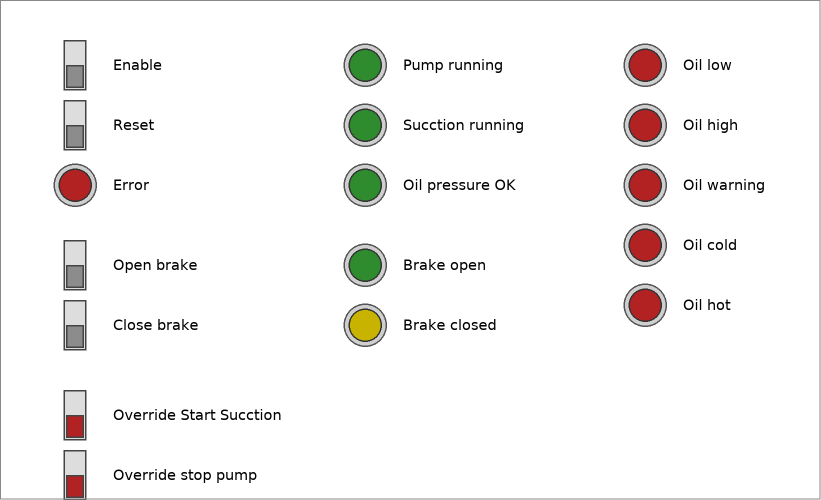
VISUALIZATION Hydraulics  // 821x500
    DipSwitch (50,40 50x50), variable: HydraulicsControl.enable, behaviour: TOGGLE, style: Switch-DipSwitch-Gray
    DipSwitch (50,100 50x50), variable: HydraulicsControl.reset, behaviour: TOGGLE, style: Switch-DipSwitch-Gray
    Label (110,50 101x30), "Enable"
    Label (110,110 101x30), "Reset"
    Lamp1 (50,160 50x50), variable: HydraulicsControl.error, style: Lamp-Lamp1-Red
    Label (110,170 101x30), "Error"
    DipSwitch (50,390 50x50), variable: HydraulicsControl.suction_manual, behaviour: TOGGLE, style: Switch-DipSwitch-Red
    DipSwitch (50,450 50x50), variable: HydraulicsControl.pump_manual_stop, behaviour: TOGGLE, style: Switch-DipSwitch-Red
    Label (110,400 171x30), "Override Start Sucction"
    Label (110,460 161x30), "Override stop pump"
    Lamp1 (340,40 50x50), variable: HydraulicsControl.pump_running, style: Lamp-Lamp1-Green
    Label (400,50 141x30), "Pump running"
    Lamp1 (340,100 50x50), variable: HydraulicsControl.suction_running, style: Lamp-Lamp1-Green
    Label (400,110 141x30), "Sucction running"
    Lamp1 (340,240 50x50), variable: HydraulicsControl.brake_open, style: Lamp-Lamp1-Green
    Label (400,250 141x30), "Brake open"
    Lamp1 (340,300 50x50), variable: HydraulicsControl.brake_closed, style: Lamp-Lamp1-Yellow
    Label (400,310 141x30), "Brake closed"
    Lamp1 (620,40 50x50), variable: HydraulicsControl.oil_low, style: Lamp-Lamp1-Red
    Label (680,50 141x30), "Oil low"
    Lamp1 (620,100 50x50), variable: HydraulicsControl.oil_high, style: Lamp-Lamp1-Red
    Label (680,110 141x30), "Oil high"
    Lamp1 (620,160 50x50), variable: HydraulicsControl.oil_warning, style: Lamp-Lamp1-Red
    Label (680,170 141x30), "Oil warning"
    Lamp1 (340,160 50x50), variable: HydraulicsControl.oil_pressure_OK, style: Lamp-Lamp1-Green
    Label (400,170 141x30), "Oil pressure OK"
    Lamp1 (620,220 50x50), variable: HydraulicsControl.oil_cold, style: Lamp-Lamp1-Red
    Label (680,230 141x30), "Oil cold"
    Lamp1 (620,280 50x50), variable: HydraulicsControl.oil_hot, style: Lamp-Lamp1-Red
    Label (680,290 141x30), "Oil hot"
    DipSwitch (50,240 50x50), variable: HydraulicsControl.iopen_brake, behaviour: TOGGLE, style: Switch-DipSwitch-Gray
    DipSwitch (50,300 50x50), variable: HydraulicsControl.iclose_brake, behaviour: TOGGLE, style: Switch-DipSwitch-Gray
    Label (110,250 101x30), "Open brake"
    Label (110,310 101x30), "Close brake"
END_VISUALIZATION

(* stored: Version 1.1.0.1, ProductVersion 3.1.4024.12
   Visu Hydraulics: Id {371113af-a8cf-42ba-8f72-dc02b3afe399} *)
